(* CODESYS project Trends.export

Project tree, tasks and I/O mapping:
  visualisation Trends
*)

// /Trends
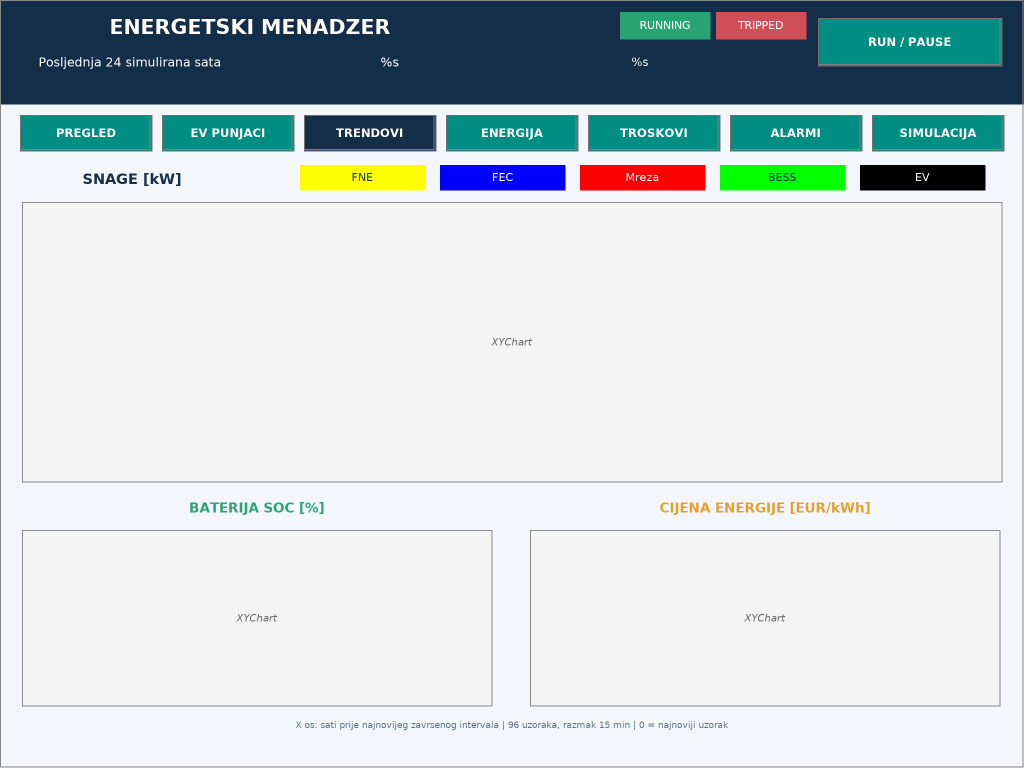
VISUALIZATION Trends  // 1024x768
    Rectangle (0,0 1024x768)
    Rectangle (0,0 1024x104)
    Rectangle (20,10 460x34), "ENERGETSKI MENADZER"
    Rectangle (20,48 220x28), "Posljednja 24 simulirana sata"
    Rectangle (260,49 260x26), "%s", text variable: Team_HMI.sDateTime
    Rectangle (530,49 220x26), "%s", text variable: Team_HMI.sPriceMode
    Button (818,18 184x48), "RUN / PAUSE"
        toggle SimCtrl.run
    Rectangle (620,12 90x27), "PAUSED", invisible if: SimCtrl.run
    Rectangle (620,12 90x27), "RUNNING", invisible if: NOT SimCtrl.run
    Rectangle (716,12 90x27), "TRIPPED", invisible if: NOT SimCtrl.tripped
    Button (20,115 132x36), "PREGLED"
        OnMouseClick:  Assign=Overview, Type=Assignment
    Button (162,115 132x36), "EV PUNJACI"
        OnMouseClick:  Assign=EVs, Type=Assignment
    Button (304,115 132x36), "TRENDOVI"
        OnMouseClick:  Assign=Trends, Type=Assignment
    Button (446,115 132x36), "ENERGIJA"
        OnMouseClick:  Assign=Energy, Type=Assignment
    Button (588,115 132x36), "TROSKOVI"
        OnMouseClick:  Assign=Costs, Type=Assignment
    Button (730,115 132x36), "ALARMI"
        OnMouseClick:  Assign=Alarms, Type=Assignment
    Button (872,115 132x36), "SIMULACIJA"
        OnMouseClick:  Assign=Controls, Type=Assignment
    Rectangle (22,165 220x28), "SNAGE [kW]"
    Rectangle (300,165 125x25), "FNE"
    Rectangle (440,165 125x25), "FEC"
    Rectangle (580,165 125x25), "Mreza"
    Rectangle (720,165 125x25), "BESS"
    Rectangle (860,165 125x25), "EV"
    XYChart (22,202 980x280)
    Rectangle (22,494 470x28), "BATERIJA SOC [%]"
    Rectangle (530,494 470x28), "CIJENA ENERGIJE [EUR/kWh]"
    XYChart (22,530 470x176)
    XYChart (530,530 470x176)
    Rectangle (22,714 980x22), "X os: sati prije najnovijeg zavrsenog intervala | 96 uzoraka, razmak 15 min | 0 = najnoviji uzorak"
END_VISUALIZATION
